// MAIN - builds the plant from HrlConfig.json, runs it in the operating mode
// the HMI asks for (eModeRequest), forced to stop while the safety interface
// does not allow motion. With mfr.link = emulator the MFR emulator drives it.
// Watch fbPlant.fbSrm (positions, jobs), fbPlant.fbRack and fbPlant.fbDiag online.
PROGRAM MAIN
VAR
    fbPlant      : FB_Hrl(ipParent := 0, sNodeName := 'HRL');
    fbOpMode     : FB_OpModeHandler;
    fbEmulator   : FB_MfrEmulator;
    fbConfig     : FB_HrlConfig;   // HrlConfig.json from the boot folder; defaults if absent
    fbHmi        : FB_HmiBridge;   // GVL_Hmi <-> plant
    eModeNow     : E_OpMode;
    bInit        : BOOL := TRUE;
END_VAR

IF bInit THEN
    fbConfig();
    IF NOT fbConfig.bDone THEN
        RETURN;   // the plant starts only with its final configuration
    END_IF
    fbPlant.stConfig     := fbConfig.stConfig;
    fbPlant.sConfigError := fbConfig.sError;
    fbOpMode.SetRoot(fbPlant);
    bInit := FALSE;
END_IF

fbHmi.Run(fbPlant, fbEmulator, GVL_Hmi.stCommand, GVL_Hmi.stStatus, eModeNow);
IF fbPlant.bSafetyOk THEN
    eModeNow := fbHmi.eModeRequest;
ELSE
    eModeNow := E_OpMode.eStop;   // safety first: no motion without the safety OK
END_IF
fbOpMode.Mode := eModeNow;
IF fbPlant.stConfig.eMfrLink = E_MfrLink.eEmulator THEN
    fbEmulator.Run(fbPlant);   // no real MFR: the emulator sends the orders
END_IF
fbOpMode.Cyclic();

END_PROGRAM

(* stored: Version 1.1.0.1
   POU MAIN: Id {b8e037f9-eaed-4553-9535-9f4c633c54c9}, SpecialFunc None *)
